FUNCTION_BLOCK Distributing_HMI (* Service Interface Function Block Type *)
  (* Standard: 61499-2 *)
  (* Version 0.0, 11/16/2026, Sandeep Patil, Flexbridge AB, template *)
  PACKAGE Flexbridge.FestoMPS400;
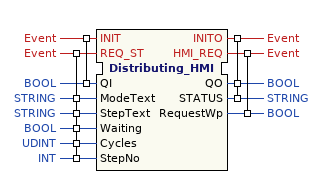
  EVENT_INPUT
    INIT WITH QI;
    REQ_ST WITH ModeText, StepText, Waiting, Cycles, StepNo;
  END_EVENT
  EVENT_OUTPUT
    INITO WITH QO, STATUS;
    HMI_REQ WITH RequestWp;
  END_EVENT
  VAR_INPUT
    QI : BOOL; (* Input event qualifier *)
    ModeText : STRING; (* Station mode *)
    StepText : STRING; (* Current step (number and name) *)
    Waiting : BOOL; (* Waiting for workpieces (magazine empty) *)
    Cycles : UDINT; (* Workpieces handed over since start-up *)
    StepNo : INT; (* Current step number *)
  END_VAR
  VAR_OUTPUT
    QO : BOOL; (* Event Output Qualifier *)
    STATUS : STRING; (* Service Status *)
    RequestWp : BOOL; (* Button: request one workpiece (stands in for Testing) *)
  END_VAR
  SERVICE /
    SEQUENCE 
    END_SEQUENCE
  END_SERVICE
END_FUNCTION_BLOCK
